Fanuc KAREL source: kt00257.KL

-- PROVISIONAL review KL for V770-1; original PC SHA256 24f98f00c3644185f4f591ac9fd1b7c04de28bb39379eeca35b1c60e119deb61
-- Incomplete behavior may be omitted. Consult companion uncertainty JSON. Do not deploy.
PROGRAM KT00257
%NOLOCKGROUP
VAR
  I1 : INTEGER
  I2 : INTEGER
  OUT : BOOLEAN
BEGIN
  -- UNRESOLVED_PC offsets 5-16; opcodes 2E,23
  -- UNRESOLVED_PC offsets 21-32; opcodes 2E,23
  -- UNRESOLVED_PC offsets 37-48; opcodes 2E,23
  -- UNRESOLVED_PC offsets 53-64; opcodes 2E,23
  -- UNRESOLVED_PC offsets 69-88; opcodes 21,21,57,23
  -- UNRESOLVED_PC offsets 93-97; opcodes 7F
END KT00257
